FUNCTION_BLOCK SortingPermissives (* Sorting-only architecture following Distribution and tutorial modules 1-4 *)
  (* Standard: 61499-2 *)
  (* Version 2.0, 2026-11-09, sorting2n, sorting2n *)
  PACKAGE Main;
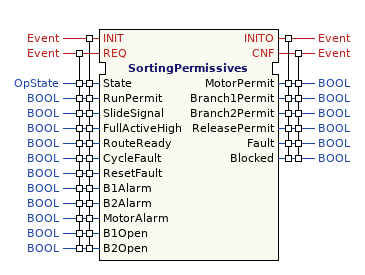
  EVENT_INPUT
    INIT WITH State, RunPermit, SlideSignal, FullActiveHigh, RouteReady, CycleFault, ResetFault, B1Alarm, B2Alarm, MotorAlarm, B1Open, B2Open;
    REQ WITH State, RunPermit, SlideSignal, FullActiveHigh, RouteReady, CycleFault, ResetFault, B1Alarm, B2Alarm, MotorAlarm, B1Open, B2Open;
  END_EVENT
  EVENT_OUTPUT
    INITO WITH MotorPermit, Branch1Permit, Branch2Permit, ReleasePermit, Fault, Blocked;
    CNF WITH MotorPermit, Branch1Permit, Branch2Permit, ReleasePermit, Fault, Blocked;
  END_EVENT
  VAR_INPUT
    State : OpState;
    RunPermit : BOOL;
    SlideSignal : BOOL;
    FullActiveHigh : BOOL;
    RouteReady : BOOL;
    CycleFault : BOOL;
    ResetFault : BOOL;
    B1Alarm : BOOL;
    B2Alarm : BOOL;
    MotorAlarm : BOOL;
    B1Open : BOOL;
    B2Open : BOOL;
  END_VAR
  VAR_OUTPUT
    MotorPermit : BOOL;
    Branch1Permit : BOOL;
    Branch2Permit : BOOL;
    ReleasePermit : BOOL;
    Fault : BOOL;
    Blocked : BOOL;
  END_VAR
  VAR
    Executing : BOOL;
  END_VAR
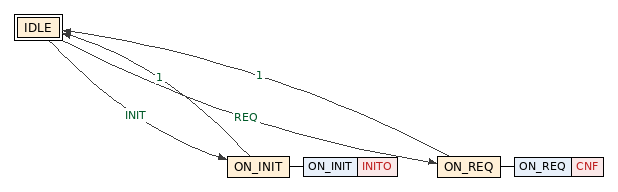
  EC_STATES
    IDLE;
    ON_INIT : ON_INIT -> INITO;
    ON_REQ : ON_REQ -> CNF;
  END_STATES
  EC_TRANSITIONS
    IDLE TO ON_INIT := INIT;
    ON_INIT TO IDLE := 1;
    IDLE TO ON_REQ := REQ;
    ON_REQ TO IDLE := 1;
  END_TRANSITIONS
  ALGORITHM ON_INIT IN ST:
IF FullActiveHigh THEN Blocked := SlideSignal; ELSE Blocked := NOT SlideSignal; END_IF;
Fault := CycleFault OR ResetFault OR B1Alarm OR B2Alarm OR MotorAlarm;
Executing := State = SE.App2StateManagement.OpState#PhaseExecute;
MotorPermit := RunPermit AND Executing AND NOT Fault;
Branch1Permit := MotorPermit AND NOT B2Open;
Branch2Permit := MotorPermit AND NOT B1Open;
ReleasePermit := MotorPermit AND RouteReady;
  END_ALGORITHM
  ALGORITHM ON_REQ IN ST:
IF FullActiveHigh THEN Blocked := SlideSignal; ELSE Blocked := NOT SlideSignal; END_IF;
Fault := CycleFault OR ResetFault OR B1Alarm OR B2Alarm OR MotorAlarm;
Executing := State = SE.App2StateManagement.OpState#PhaseExecute;
MotorPermit := RunPermit AND Executing AND NOT Fault;
Branch1Permit := MotorPermit AND NOT B2Open;
Branch2Permit := MotorPermit AND NOT B1Open;
ReleasePermit := MotorPermit AND RouteReady;
  END_ALGORITHM
END_FUNCTION_BLOCK
